(* IEC 61131-3 sources: llm-plc-st-eval/data/processed_definitivo/claude-sonnet-4-6/C4/few_shot, 3 files *)

(* ---- ejec_1.st ---- *)
FUNCTION_BLOCK FB_D
VAR_INPUT
    demanda : BOOL;  (* Señal de solicitud de caudal/presión *)
    falla1  : BOOL;  (* Fallo detectado en bomba 1 (p.ej. térmico, caudal) *)
    falla2  : BOOL;  (* Fallo detectado en bomba 2 *)
END_VAR
VAR_OUTPUT
    bomba1   : BOOL; (* Orden de marcha a bomba 1 *)
    bomba2   : BOOL; (* Orden de marcha a bomba 2 *)
    almFalla : BOOL; (* Alarma activa: la bomba de turno ha fallado *)
END_VAR
VAR
    turno : BOOL;   (* FALSE = turno de bomba 2 prioritaria,
                       TRUE  = turno de bomba 1 prioritaria *)
    fDem  : R_TRIG; (* Detector de flanco ascendente sobre 'demanda' *)
END_VAR

(* ── Detección de flanco ascendente de demanda ──────────────────────────
   fDem.Q vale TRUE únicamente durante el ciclo en que 'demanda'
   pasa de FALSE a TRUE; se usa para alternar el turno en cada
   nueva solicitud, no en cada ciclo de scan.                          *)
fDem(CLK := demanda);

(* ── Alternancia de turno ───────────────────────────────────────────────
   Con cada nuevo flanco de demanda se invierte la bomba prioritaria,
   distribuyendo las horas de funcionamiento entre ambas unidades.     *)
IF fDem.Q THEN
    turno := NOT turno;
END_IF

(* ── Lógica de arranque con redundancia ─────────────────────────────── *)
IF demanda THEN

    IF turno THEN
        (* Turno de bomba 1 como unidad principal *)
        bomba1 := NOT falla1;              (* Arranca bomba 1 si no falla *)
        bomba2 := falla1 AND NOT falla2;   (* Bomba 2 entra solo si bomba 1 falla
                                              y bomba 2 está sana              *)
        almFalla := falla1;                (* Alarma si la unidad prioritaria falla *)

    ELSE
        (* Turno de bomba 2 como unidad principal *)
        bomba2 := NOT falla2;              (* Arranca bomba 2 si no falla *)
        bomba1 := falla2 AND NOT falla1;   (* Bomba 1 entra solo si bomba 2 falla
                                              y bomba 1 está sana              *)
        almFalla := falla2;                (* Alarma si la unidad prioritaria falla *)
    END_IF

ELSE
    (* ── Sin demanda: apagado total y reset de alarma ───────────────── *)
    bomba1   := FALSE;
    bomba2   := FALSE;
    almFalla := FALSE;
END_IF

END_FUNCTION_BLOCK

(* ---- ejec_2.st ---- *)
FUNCTION_BLOCK FB_D
VAR_INPUT
    demanda : BOOL;  (* Señal de demanda de caudal: TRUE = se requiere bombeo *)
    falla1  : BOOL;  (* Fallo detectado en bomba 1: TRUE = bomba 1 en falla *)
    falla2  : BOOL;  (* Fallo detectado en bomba 2: TRUE = bomba 2 en falla *)
END_VAR
VAR_OUTPUT
    bomba1   : BOOL; (* Orden de marcha a bomba 1 *)
    bomba2   : BOOL; (* Orden de marcha a bomba 2 *)
    almFalla : BOOL; (* Alarma activa: la bomba de turno tiene falla *)
END_VAR
VAR
    turno : BOOL;   (* Bit de alternancia: FALSE = turno de bomba 2, TRUE = turno de bomba 1 *)
    fDem  : R_TRIG; (* Detector de flanco ascendente sobre la señal de demanda *)
END_VAR

(* ── Detección de flanco ascendente de demanda ──────────────────────────────
   fDem.Q vale TRUE únicamente durante el ciclo en que demanda pasa de 0 a 1. *)
fDem(CLK := demanda);

(* ── Alternancia de turno ────────────────────────────────────────────────────
   Cada nuevo arranque (flanco de demanda) invierte el bit de turno,
   asegurando que las bombas se usen de forma alternada y equitativa. *)
IF fDem.Q THEN
    turno := NOT turno;
END_IF

(* ── Lógica de arranque y alarma ─────────────────────────────────────────── *)
IF demanda THEN

    IF turno THEN
        (* Turno de bomba 1 como unidad prioritaria *)
        bomba1   := NOT falla1;          (* Arranca bomba 1 si no tiene falla *)
        bomba2   := falla1 AND NOT falla2; (* Bomba 2 entra solo si bomba 1 falla y bomba 2 está sana *)
        almFalla := falla1;              (* Alarma si la unidad prioritaria (bomba 1) está en falla *)
    ELSE
        (* Turno de bomba 2 como unidad prioritaria *)
        bomba2   := NOT falla2;          (* Arranca bomba 2 si no tiene falla *)
        bomba1   := falla2 AND NOT falla1; (* Bomba 1 entra solo si bomba 2 falla y bomba 1 está sana *)
        almFalla := falla2;              (* Alarma si la unidad prioritaria (bomba 2) está en falla *)
    END_IF

ELSE
    (* Sin demanda: apagado total y alarma silenciada *)
    bomba1   := FALSE;
    bomba2   := FALSE;
    almFalla := FALSE;
END_IF

END_FUNCTION_BLOCK

(* ---- ejec_3.st ---- *)
FUNCTION_BLOCK FB_D
VAR_INPUT
    demanda : BOOL;  (* Señal de solicitud de bombeo (TRUE = se requiere caudal) *)
    falla1  : BOOL;  (* Señal de falla de la bomba 1 (TRUE = bomba 1 en falla) *)
    falla2  : BOOL;  (* Señal de falla de la bomba 2 (TRUE = bomba 2 en falla) *)
END_VAR
VAR_OUTPUT
    bomba1   : BOOL; (* Comando de arranque de la bomba 1 *)
    bomba2   : BOOL; (* Comando de arranque de la bomba 2 *)
    almFalla : BOOL; (* Alarma activa cuando la bomba prioritaria está en falla *)
END_VAR
VAR
    turno : BOOL;   (* FALSE = turno de bomba 2 como prioritaria;
                       TRUE  = turno de bomba 1 como prioritaria *)
    fDem  : R_TRIG; (* Detector de flanco ascendente sobre la señal de demanda *)
END_VAR

(* ── Detección de flanco ascendente de demanda ───────────────────────────────
   Cada vez que demanda pasa de FALSE a TRUE se genera un pulso en fDem.Q.
   Esto permite alternar el turno exactamente una vez por cada nueva solicitud. *)
fDem(CLK := demanda);

(* ── Alternancia de turno ────────────────────────────────────────────────────
   En cada flanco ascendente de demanda se invierte la variable turno,
   cambiando qué bomba actúa como prioritaria en el siguiente ciclo de bombeo. *)
IF fDem.Q THEN
    turno := NOT turno;
END_IF

(* ── Lógica de arranque y respaldo ───────────────────────────────────────────
   Solo se activan bombas mientras la demanda esté presente. *)
IF demanda THEN

    (* ── Turno de bomba 1 como prioritaria ───────────────────────────────── *)
    IF turno THEN
        (* Bomba 1 arranca si no tiene falla propia *)
        bomba1 := NOT falla1;

        (* Bomba 2 entra como respaldo únicamente si bomba 1 falló
           y ella misma no presenta falla *)
        bomba2 := falla1 AND NOT falla2;

        (* Alarma activa si la bomba prioritaria (bomba 1) está en falla *)
        almFalla := falla1;

    (* ── Turno de bomba 2 como prioritaria ───────────────────────────────── *)
    ELSE
        (* Bomba 2 arranca si no tiene falla propia *)
        bomba2 := NOT falla2;

        (* Bomba 1 entra como respaldo únicamente si bomba 2 falló
           y ella misma no presenta falla *)
        bomba1 := falla2 AND NOT falla1;

        (* Alarma activa si la bomba prioritaria (bomba 2) está en falla *)
        almFalla := falla2;
    END_IF

(* ── Sin demanda: todo apagado ───────────────────────────────────────────────
   Se fuerzan a FALSE todas las salidas para garantizar estado seguro
   cuando no se requiere bombeo. *)
ELSE
    bomba1   := FALSE;
    bomba2   := FALSE;
    almFalla := FALSE;
END_IF

END_FUNCTION_BLOCK
